// TIA Portal V20 export
Screen "200RB04_Stand_V23"  1276x673
  ScreenItem "Line_Header_X0_Y64" at 0,64 size 1276x0  Type=HmiLine
  ScreenItem "permanentareaborderrectangle" at 0,0 size 0x0  Type=HmiRectangle
  ScreenItem "Button_Back" at 2,2 size 90x60  Type=HmiButton
  ScreenItem "Title_ScreenOverview_X390_Y2_1" at 390,3 size 510x57  Type=HmiTextBox
  ScreenItem "Title_ScreenOverview_X390_Y2_5" at 1130,78 size 139x57  Type=HmiTextBox
  ScreenItem "Title_ScreenOverview_X390_Y2_6" at 1130,144 size 139x57  Type=HmiTextBox
  ScreenItem "Title_ScreenOverview_X390_Y2_7" at 1130,144 size 139x57  Type=HmiTextBox
  ScreenItem "Graphic view_1" at 457,157 size 358x495  Type=HmiGraphicView
  ScreenItem "Line_7" at 745,243 size 76x1  Type=HmiLine
  ScreenItem "Line_1" at 433,150 size 136x59  Type=HmiLine
  ScreenItem "Line_2" at 703,151 size 112x60  Type=HmiLine
  ScreenItem "Rectangle_3" at 0,0 size 166x43  Type=HmiRectangle
  ScreenItem "文本域_3" at 2,1 size 134x40  Type=HmiTextBox
  ScreenItem "圆_3" at 0,0 size 100x30  Type=HmiCircle
  ScreenItem "圆_4" at 0,0 size 100x30  Type=HmiCircle
  ScreenItem "Rectangle_1" at 0,0 size 166x43  Type=HmiRectangle
  ScreenItem "文本域_1" at 2,1 size 134x40  Type=HmiTextBox
  ScreenItem "圆_1" at 0,0 size 100x30  Type=HmiCircle
  ScreenItem "圆_2" at 0,0 size 100x30  Type=HmiCircle
  ScreenItem "Rectangle_9" at 855,263 size 52x43  Type=HmiRectangle
  ScreenItem "文本域_9" at 814,220 size 134x40  Type=HmiTextBox
  ScreenItem "Title_ScreenOverview_X390_Y2_17" at 855,284 size 25x21  Type=HmiTextBox
  ScreenItem "Title_ScreenOverview_X390_Y2_18" at 882,284 size 25x21  Type=HmiTextBox
  ScreenItem "Title_ScreenOverview_X390_Y2_19" at 855,264 size 52x19  Type=HmiTextBox
